// TIA Portal V20 export
DATA_BLOCK "DB_Manual"   // DB8
{ S7_Optimized_Access := 'TRUE' }
// stored: MemoryReserve 100
   VAR
      xManEtiketa : Bool;   // TRUE = světla + trigger etiketa
      xManFolie : Bool;   // TRUE = světla + trigger folie
      test_vyr : Bool;
   END_VAR
BEGIN
END_DATA_BLOCK
